Fanuc KAREL source: KT00868.KL

PROGRAM KT00868
%NOLOCKGROUP
VAR
  I1: INTEGER
  I2: INTEGER
  OUT: INTEGER
BEGIN
  I1 = 2
  I2 = 3
  I1 = 2
  I2 = 3
  OUT = TRUNC(I1)
END KT00868
